(* IEC 61131-3 sources: STAR-PLC-Agent/results/raw/four_group_20261114/star_deepseek_v4/PUB018/generation/sim_00, 1 file *)

(* ---- test_program.st ---- *)
PROGRAM PLC_PRG
VAR
 BenchStep : UDINT := 0;
 BenchCalls : UDINT := 0;
 BenchDone : BOOL := FALSE;
 BenchUut0 : FB_Task;
 BenchUut1 : FB_Task;
 Binding_0_item : DINT;
 Binding_0_buffer : DINT;
 Binding_1_item : DINT;
 Binding_1_buffer : DINT;
 TraceIn_enqueue : ARRAY[0..15] OF BOOL;
 TraceIn_dequeue : ARRAY[0..15] OF BOOL;
 TraceIn_reset : ARRAY[0..15] OF BOOL;
 TraceOut_elementCount : ARRAY[0..15] OF DINT;
 TraceOut_status : ARRAY[0..15] OF WORD;
 TraceOut_item_DINT : ARRAY[0..15] OF DINT;
 TraceOut_item_BOOL : ARRAY[0..15] OF BOOL;
 TraceInIO_item_DINT : ARRAY[0..15] OF DINT;
END_VAR

IF NOT BenchDone THEN
 CASE BenchStep OF
 0:
   Binding_0_item := DINT#0;
   BenchUut0.enqueue := FALSE;
   BenchUut0.dequeue := FALSE;
   BenchUut0.reset := FALSE;
   TraceIn_enqueue[0] := BenchUut0.enqueue;
   TraceIn_dequeue[0] := BenchUut0.dequeue;
   TraceIn_reset[0] := BenchUut0.reset;
   TraceInIO_item_DINT[0] := Binding_0_item;
   BenchUut0(item := Binding_0_item, buffer := Binding_0_buffer);
   TraceOut_elementCount[0] := BenchUut0.elementCount;
   TraceOut_status[0] := BenchUut0.status;
   TraceOut_item_DINT[0] := Binding_0_item;
   BenchCalls := BenchCalls + 1;
 1:
   Binding_0_item := DINT#11;
   BenchUut0.enqueue := TRUE;
   BenchUut0.dequeue := FALSE;
   BenchUut0.reset := FALSE;
   TraceIn_enqueue[1] := BenchUut0.enqueue;
   TraceIn_dequeue[1] := BenchUut0.dequeue;
   TraceIn_reset[1] := BenchUut0.reset;
   TraceInIO_item_DINT[1] := Binding_0_item;
   BenchUut0(item := Binding_0_item, buffer := Binding_0_buffer);
   TraceOut_elementCount[1] := BenchUut0.elementCount;
   TraceOut_status[1] := BenchUut0.status;
   TraceOut_item_DINT[1] := Binding_0_item;
   BenchCalls := BenchCalls + 1;
 2:
   Binding_0_item := DINT#12;
   BenchUut0.enqueue := FALSE;
   BenchUut0.dequeue := FALSE;
   BenchUut0.reset := FALSE;
   TraceIn_enqueue[2] := BenchUut0.enqueue;
   TraceIn_dequeue[2] := BenchUut0.dequeue;
   TraceIn_reset[2] := BenchUut0.reset;
   TraceInIO_item_DINT[2] := Binding_0_item;
   BenchUut0(item := Binding_0_item, buffer := Binding_0_buffer);
   TraceOut_elementCount[2] := BenchUut0.elementCount;
   TraceOut_status[2] := BenchUut0.status;
   TraceOut_item_DINT[2] := Binding_0_item;
   BenchCalls := BenchCalls + 1;
 3:
   Binding_0_item := DINT#22;
   BenchUut0.enqueue := TRUE;
   BenchUut0.dequeue := FALSE;
   BenchUut0.reset := FALSE;
   TraceIn_enqueue[3] := BenchUut0.enqueue;
   TraceIn_dequeue[3] := BenchUut0.dequeue;
   TraceIn_reset[3] := BenchUut0.reset;
   TraceInIO_item_DINT[3] := Binding_0_item;
   BenchUut0(item := Binding_0_item, buffer := Binding_0_buffer);
   TraceOut_elementCount[3] := BenchUut0.elementCount;
   TraceOut_status[3] := BenchUut0.status;
   TraceOut_item_DINT[3] := Binding_0_item;
   BenchCalls := BenchCalls + 1;
 4:
   Binding_0_item := DINT#0;
   BenchUut0.enqueue := FALSE;
   BenchUut0.dequeue := TRUE;
   BenchUut0.reset := FALSE;
   TraceIn_enqueue[4] := BenchUut0.enqueue;
   TraceIn_dequeue[4] := BenchUut0.dequeue;
   TraceIn_reset[4] := BenchUut0.reset;
   TraceInIO_item_DINT[4] := Binding_0_item;
   BenchUut0(item := Binding_0_item, buffer := Binding_0_buffer);
   TraceOut_elementCount[4] := BenchUut0.elementCount;
   TraceOut_status[4] := BenchUut0.status;
   TraceOut_item_DINT[4] := Binding_0_item;
   BenchCalls := BenchCalls + 1;
 5:
   Binding_0_item := DINT#33;
   BenchUut0.enqueue := TRUE;
   BenchUut0.dequeue := FALSE;
   BenchUut0.reset := FALSE;
   TraceIn_enqueue[5] := BenchUut0.enqueue;
   TraceIn_dequeue[5] := BenchUut0.dequeue;
   TraceIn_reset[5] := BenchUut0.reset;
   TraceInIO_item_DINT[5] := Binding_0_item;
   BenchUut0(item := Binding_0_item, buffer := Binding_0_buffer);
   TraceOut_elementCount[5] := BenchUut0.elementCount;
   TraceOut_status[5] := BenchUut0.status;
   TraceOut_item_DINT[5] := Binding_0_item;
   BenchCalls := BenchCalls + 1;
 6:
   Binding_0_item := DINT#0;
   BenchUut0.enqueue := FALSE;
   BenchUut0.dequeue := FALSE;
   BenchUut0.reset := FALSE;
   TraceIn_enqueue[6] := BenchUut0.enqueue;
   TraceIn_dequeue[6] := BenchUut0.dequeue;
   TraceIn_reset[6] := BenchUut0.reset;
   TraceInIO_item_DINT[6] := Binding_0_item;
   BenchUut0(item := Binding_0_item, buffer := Binding_0_buffer);
   TraceOut_elementCount[6] := BenchUut0.elementCount;
   TraceOut_status[6] := BenchUut0.status;
   TraceOut_item_DINT[6] := Binding_0_item;
   BenchCalls := BenchCalls + 1;
 7:
   Binding_0_item := DINT#0;
   BenchUut0.enqueue := FALSE;
   BenchUut0.dequeue := TRUE;
   BenchUut0.reset := FALSE;
   TraceIn_enqueue[7] := BenchUut0.enqueue;
   TraceIn_dequeue[7] := BenchUut0.dequeue;
   TraceIn_reset[7] := BenchUut0.reset;
   TraceInIO_item_DINT[7] := Binding_0_item;
   BenchUut0(item := Binding_0_item, buffer := Binding_0_buffer);
   TraceOut_elementCount[7] := BenchUut0.elementCount;
   TraceOut_status[7] := BenchUut0.status;
   TraceOut_item_DINT[7] := Binding_0_item;
   BenchCalls := BenchCalls + 1;
 8:
   Binding_1_item := DINT#0;
   BenchUut1.enqueue := FALSE;
   BenchUut1.dequeue := FALSE;
   BenchUut1.reset := FALSE;
   TraceIn_enqueue[8] := BenchUut1.enqueue;
   TraceIn_dequeue[8] := BenchUut1.dequeue;
   TraceIn_reset[8] := BenchUut1.reset;
   TraceInIO_item_DINT[8] := Binding_1_item;
   BenchUut1(item := Binding_1_item, buffer := Binding_1_buffer);
   TraceOut_elementCount[8] := BenchUut1.elementCount;
   TraceOut_status[8] := BenchUut1.status;
   TraceOut_item_DINT[8] := Binding_1_item;
   BenchCalls := BenchCalls + 1;
 9:
   Binding_1_item := DINT#5;
   BenchUut1.enqueue := FALSE;
   BenchUut1.dequeue := TRUE;
   BenchUut1.reset := FALSE;
   TraceIn_enqueue[9] := BenchUut1.enqueue;
   TraceIn_dequeue[9] := BenchUut1.dequeue;
   TraceIn_reset[9] := BenchUut1.reset;
   TraceInIO_item_DINT[9] := Binding_1_item;
   BenchUut1(item := Binding_1_item, buffer := Binding_1_buffer);
   TraceOut_elementCount[9] := BenchUut1.elementCount;
   TraceOut_status[9] := BenchUut1.status;
   TraceOut_item_DINT[9] := Binding_1_item;
   BenchCalls := BenchCalls + 1;
 10:
   Binding_1_item := DINT#11;
   BenchUut1.enqueue := TRUE;
   BenchUut1.dequeue := FALSE;
   BenchUut1.reset := FALSE;
   TraceIn_enqueue[10] := BenchUut1.enqueue;
   TraceIn_dequeue[10] := BenchUut1.dequeue;
   TraceIn_reset[10] := BenchUut1.reset;
   TraceInIO_item_DINT[10] := Binding_1_item;
   BenchUut1(item := Binding_1_item, buffer := Binding_1_buffer);
   TraceOut_elementCount[10] := BenchUut1.elementCount;
   TraceOut_status[10] := BenchUut1.status;
   TraceOut_item_DINT[10] := Binding_1_item;
   BenchCalls := BenchCalls + 1;
 11:
   Binding_1_item := DINT#12;
   BenchUut1.enqueue := FALSE;
   BenchUut1.dequeue := FALSE;
   BenchUut1.reset := FALSE;
   TraceIn_enqueue[11] := BenchUut1.enqueue;
   TraceIn_dequeue[11] := BenchUut1.dequeue;
   TraceIn_reset[11] := BenchUut1.reset;
   TraceInIO_item_DINT[11] := Binding_1_item;
   BenchUut1(item := Binding_1_item, buffer := Binding_1_buffer);
   TraceOut_elementCount[11] := BenchUut1.elementCount;
   TraceOut_status[11] := BenchUut1.status;
   TraceOut_item_DINT[11] := Binding_1_item;
   BenchCalls := BenchCalls + 1;
 12:
   Binding_1_item := DINT#22;
   BenchUut1.enqueue := TRUE;
   BenchUut1.dequeue := FALSE;
   BenchUut1.reset := FALSE;
   TraceIn_enqueue[12] := BenchUut1.enqueue;
   TraceIn_dequeue[12] := BenchUut1.dequeue;
   TraceIn_reset[12] := BenchUut1.reset;
   TraceInIO_item_DINT[12] := Binding_1_item;
   BenchUut1(item := Binding_1_item, buffer := Binding_1_buffer);
   TraceOut_elementCount[12] := BenchUut1.elementCount;
   TraceOut_status[12] := BenchUut1.status;
   TraceOut_item_DINT[12] := Binding_1_item;
   BenchCalls := BenchCalls + 1;
 13:
   Binding_1_item := DINT#33;
   BenchUut1.enqueue := FALSE;
   BenchUut1.dequeue := FALSE;
   BenchUut1.reset := FALSE;
   TraceIn_enqueue[13] := BenchUut1.enqueue;
   TraceIn_dequeue[13] := BenchUut1.dequeue;
   TraceIn_reset[13] := BenchUut1.reset;
   TraceInIO_item_DINT[13] := Binding_1_item;
   BenchUut1(item := Binding_1_item, buffer := Binding_1_buffer);
   TraceOut_elementCount[13] := BenchUut1.elementCount;
   TraceOut_status[13] := BenchUut1.status;
   TraceOut_item_DINT[13] := Binding_1_item;
   BenchCalls := BenchCalls + 1;
 14:
   Binding_1_item := DINT#33;
   BenchUut1.enqueue := TRUE;
   BenchUut1.dequeue := FALSE;
   BenchUut1.reset := FALSE;
   TraceIn_enqueue[14] := BenchUut1.enqueue;
   TraceIn_dequeue[14] := BenchUut1.dequeue;
   TraceIn_reset[14] := BenchUut1.reset;
   TraceInIO_item_DINT[14] := Binding_1_item;
   BenchUut1(item := Binding_1_item, buffer := Binding_1_buffer);
   TraceOut_elementCount[14] := BenchUut1.elementCount;
   TraceOut_status[14] := BenchUut1.status;
   TraceOut_item_DINT[14] := Binding_1_item;
   BenchCalls := BenchCalls + 1;
 15:
   Binding_1_item := DINT#99;
   BenchUut1.enqueue := FALSE;
   BenchUut1.dequeue := TRUE;
   BenchUut1.reset := TRUE;
   TraceIn_enqueue[15] := BenchUut1.enqueue;
   TraceIn_dequeue[15] := BenchUut1.dequeue;
   TraceIn_reset[15] := BenchUut1.reset;
   TraceInIO_item_DINT[15] := Binding_1_item;
   BenchUut1(item := Binding_1_item, buffer := Binding_1_buffer);
   TraceOut_elementCount[15] := BenchUut1.elementCount;
   TraceOut_status[15] := BenchUut1.status;
   TraceOut_item_DINT[15] := Binding_1_item;
   BenchCalls := BenchCalls + 1;
 END_CASE;
 BenchStep := BenchStep + 1;
 IF BenchStep >= 16 THEN BenchDone := TRUE; END_IF;
END_IF;
END_PROGRAM
